// TIA Portal V20 export
// export: Created 2026-10-19T18:37:09.630453Z, ExportSetting WithDefaults, DisplayName Totally Integrated Automation Portal, DisplayVersion V20 Update 6, DisplayName TIA Portal Openness, DisplayVersion V20 Update 6, DisplayName TIA Portal Version Control Interface, DisplayVersion V20 Update 6, DisplayName SINAMICS Startdrive Advanced, DisplayVersion V20 SP1, DisplayName SINAMICS Startdrive G130, G150, S120, S150, SINAMICS MV, G220, S200, S210, DisplayVersion V20 SP1, DisplayName SINAMICS Startdrive G110M, G120, G120C, G120D, G120P, G115D, DisplayVersion V20 SP1, DisplayName STEP 7 Professional, DisplayVersion V20 Update 6, DisplayName STEP 7 Safety, DisplayVersion V20 Update 2, DisplayName WinCC Basic/Comfort/Advanced, DisplayVersion V20 Update 6, DisplayName WinCC Unified, DisplayVersion V20 Update 6
FUNCTION_BLOCK "VTD_HMI_FB"   // FB14, SCL
{ S7_Optimized_Access := 'TRUE' }
VERSION : 0.1
// stored: AutoNumber true, IsIECCheckEnabled false, IsRetainMemResEnabled false, MemoryReserve 100, SetENOAutomatically false, UDAEnableTagReadback false
   VAR
      T_Charge { S7_SetPoint := 'True'} : TON_TIME;
   END_VAR
BEGIN
   //CHARGE DATA CHANGING CONVEYORS ID
   IF "VTD_System_Selected_HMI" <> "VTD_ID_HMI_OLD" THEN
       "Screen_DB".Charge_VTD_Commands := TRUE;
       "VTD_ID_HMI_OLD" := "VTD_System_Selected_HMI";
   END_IF;

   //CHARGE ONCE THE COMMANDS STATUS
   IF "Screen_DB".Charge_VTD_Commands THEN
       CASE "VTD_System_Selected_HMI" OF
           1:
               "VTD_Mode_Change_HMI" := "Control_DB".VTD_Sys[1].Mode;
               "VTD_Enable_HMI" := "Control_DB".VTD_Sys[1].Instruction.Enable;
               "LE_Bypass" := "LE_Bypass(1)";
               "VTD_Stop_HMI" := "Control_DB".VTD_Sys[1].Instruction.Stop;
           2:
               "VTD_Mode_Change_HMI" := "Control_DB".VTD_Sys[2].Mode;
               "VTD_Enable_HMI" := "Control_DB".VTD_Sys[2].Instruction.Enable;
               "LE_Bypass" := "LE_Bypass(2)";
               "VTD_Stop_HMI" := "Control_DB".VTD_Sys[2].Instruction.Stop;
       END_CASE;

       #T_Charge.TON(IN := TRUE,
                     PT := T#500mS);
       IF #T_Charge.Q THEN
           #T_Charge.TON(IN := FALSE,
                         PT := T#0mS);
           "Screen_DB".Charge_VTD_Commands := 0;
       END_IF;

   // CHARGE DATA FROM HMI (AFTER CHARGE DATA)
   ELSIF "HMI_DB".ScreenNo_Main = 1 AND NOT "Screen_DB".Charge_VTD_Commands THEN
       CASE "VTD_System_Selected_HMI" OF
           1:
               "Feed_VTD_HMI_FC"(Sys_No := 1,
                                 Rem_Loc_Keys:= "HMI_DB".Rem_Loc_Keys[1].Level,
                                 Safety_OK := "Remote_Panel_DB_1".Safety_OK,
                                 BCD_Test_Ok_HMI := "SICK_Lector_DB_1".Test_OK,
                                 BCD_Error_HMI := "SICK_Lector_DB_1".Error,
                                 BCD_RdDone := "SICK_Lector_DB_1".RdDone,
                                 BCD_ReqDone := "SICK_Lector_DB_1".ReqDone,
                                 BCD_ReqBusy := "SICK_Lector_DB_1".ReqBusy,
                                 Start_InBarcodeStation := "Start_InBarcodeStation_HMI",
                                 Sick_Lector_Reseult := "SICK_Lector_DB_1".Barcode_Result,
                                 Level_Below_Extractor := "VTD_FB_DB_1".LevelBelowExtractor,
                                 Speed_mm_s := "VTD_FB_DB_1".VTDSpeed_mm_s,
                                 LE_Bypass := "LE_Bypass(1)",
                                 BCD_Start_Comm_Test_HMI := "BCD_Test_Comm_HMI(1)",
                                 BCD_Enable_Trigger_HMI := "BCD_Enable_Trigger_HMI(1)",
                                 BCD_Disable_Trigger_HMI := "BCD_Disable_Trigger_HMI(1)",
                                 BCD_Execute_Function := "SICK_Lector_Control_DB_1".Enable_Req,
                                 System_Busy => "System_1_Busy");

           2:
               "Feed_VTD_HMI_FC"(Sys_No := 2,
                                 Rem_Loc_Keys:="HMI_DB".Rem_Loc_Keys[2].Level,
                                 Safety_OK := "Remote_Panel_DB_2".Safety_OK,
                                 BCD_Test_Ok_HMI := "SICK_Lector_DB_2".Test_OK,
                                 BCD_Error_HMI := "SICK_Lector_DB_2".Error,
                                 BCD_RdDone := "SICK_Lector_DB_2".RdDone,
                                 BCD_ReqDone := "SICK_Lector_DB_2".ReqDone,
                                 BCD_ReqBusy := "SICK_Lector_DB_2".ReqBusy,
                                 Start_InBarcodeStation := "Start_InBarcodeStation_HMI",
                                 Sick_Lector_Reseult := "SICK_Lector_DB_2".Barcode_Result,
                                 Level_Below_Extractor := "VTD_FB_DB_2".LevelBelowExtractor,
                                 Speed_mm_s := "VTD_FB_DB_2".VTDSpeed_mm_s,
                                 LE_Bypass := "LE_Bypass(2)",
                                 BCD_Start_Comm_Test_HMI := "BCD_Test_Comm_HMI(2)",
                                 BCD_Enable_Trigger_HMI := "BCD_Enable_Trigger_HMI(2)",
                                 BCD_Disable_Trigger_HMI := "BCD_Disable_Trigger_HMI(2)",
                                 BCD_Execute_Function := "SICK_Lector_Control_DB_2".Enable_Req,
                                 System_Busy => "System_2_Busy");
       END_CASE;
   END_IF;
END_FUNCTION_BLOCK
